(* PLC project Vn_int_literal_assign, Beckhoff Automation GmbH TwinCAT PLC Control 3.5.13.21 *)
(* stored: creationDateTime 1970-01-01T00:00:00 *)

PROGRAM Vn_int_literal_assign

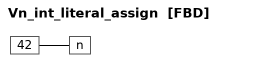
(* FBD diagram, written out as Structured Text *)
n := 42;
END_PROGRAM
